// TIA Portal V21 export
// export: Created 2026-10-12T11:32:13.9780847Z, ExportSetting WithDefaults, DisplayName Totally Integrated Automation Portal, DisplayVersion V21, DisplayName STEP 7 Professional, DisplayVersion V21, DisplayName STEP 7 Safety, DisplayVersion V21, DisplayName Tech WebApplication, DisplayVersion V21, DisplayName WinCC Basic/Comfort/Advanced, DisplayVersion V21, DisplayName WinCC Unified, DisplayVersion V21
DATA_BLOCK "DB_HMI"   // DB1
{ S7_Optimized_Access := 'FALSE' }
VERSION : 0.1
// stored: AutoNumber true, DBAccessibleFromOPCUA true, IsOnlyStoredInLoadMemory false, IsWriteProtectedInAS false
   VAR RETAIN
      "FAULT RESET PB" : Bool;
      "MOTOR JOG FWD PB" : Bool;
      "MOTOR JOG REV PB" : Bool;
      "STOP TIME" : DInt;
      "CAMERA DONE" : Bool;
   END_VAR
BEGIN
END_DATA_BLOCK
